TYPE ST_FastRefereneValueFROMPLC :
STRUCT
	(* Fast Referene Value *)
	nOverride					:INT;			(* Value of override 16384 = 100 %. *)
	nSpeed						:INT;			(* Relative speed reference value *)
	bHWLimitMax					:BOOL;			(* Hardware limit switch maximum end of range *)
	bHWLimitMin					:BOOL;			(* Hardware limit switch minimum end of range *)
END_STRUCT
END_TYPE

(* stored: Version 1.1.0.1, ProductVersion 3.1.4024.15
   DUT ST_FastRefereneValueFROMPLC: Id {f45c3c77-33ef-48d4-850b-eb6a5813b83a} *)
